Fanuc KAREL source: kc00010.KL

-- PROVISIONAL review KL for V1013-1; original PC SHA256 cbd98760c7a37dede632508e5e31ba2f387584c0e3e1743291c8938f042b91c5
-- Incomplete behavior may be omitted. Consult companion uncertainty JSON. Do not deploy.
PROGRAM KC00010
%NOLOCKGROUP
BEGIN
  -- UNRESOLVED_PC offsets 5-27; opcodes 27,22,1C,31,23
  -- UNRESOLVED_PC offsets 32-36; opcodes 7F
END KC00010
